// Mitsubishi GX Works2 project: Task2_Ex_2   PLC: FX3G

PROGRAM MAIN
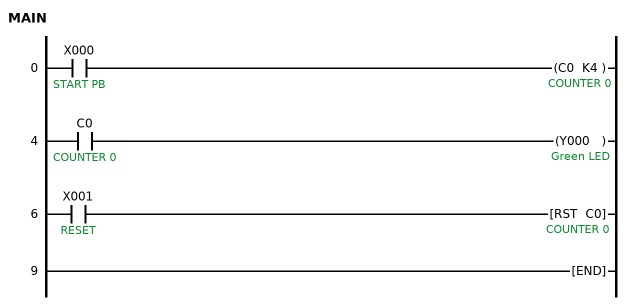
0     LD      X000  ; START PB
      OUT     C0 K4  ; COUNTER 0
4     LD      C0  ; COUNTER 0
      OUT     Y000  ; Green LED
6     LD      X001  ; RESET
      RST     C0  ; COUNTER 0
9     END
END_PROGRAM
